(* PLC project sfc_elevator_door_bomb, Anonymous Benchmark Suite 1.0 *)
(* stored: creationDateTime 2026-08-26T00:00:00 *)

PROGRAM car_control
  VAR_INPUT
    call : BOOL;
    dwell_done : BOOL;
    door_closed : BOOL;
    at_floor : BOOL;
  END_VAR
  VAR_OUTPUT
    door_open : BOOL;
    moving : BOOL;
  END_VAR

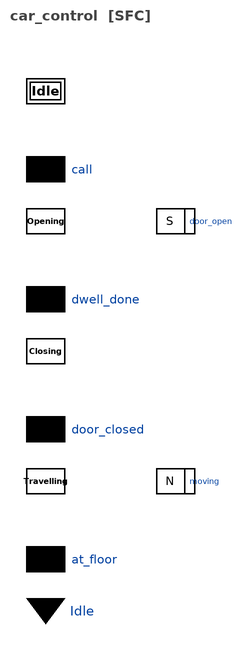
INITIAL_STEP Idle:
END_STEP
TRANSITION FROM Idle TO Opening
  := call;
END_TRANSITION
STEP Opening:
  door_open(S);
END_STEP
TRANSITION FROM Opening TO Closing
  := dwell_done;
END_TRANSITION
STEP Closing:
END_STEP
TRANSITION FROM Closing TO Travelling
  := door_closed;
END_TRANSITION
STEP Travelling:
  moving(N);
END_STEP
TRANSITION FROM Travelling TO Idle
  := at_floor;
END_TRANSITION
END_PROGRAM

CONFIGURATION Config0
  RESOURCE Res0 ON PLC
    TASK tcyclic(INTERVAL := T#10ms, PRIORITY := 0);
    PROGRAM inst0 WITH tcyclic : car_control;
  END_RESOURCE
END_CONFIGURATION
